SUBAPPLICATION Uebung_142_AX (* Übung zu NMEA 2000 Fast Packet senden (PGN 0x1FF00, 32 Byte) *)
  (* Standard: 61499-2; Description: Copyright (c) 2026 Meisterschulen am Ostbahnhof This program and the accompanying materials are made available under the terms of the Eclipse Public License 2.0 which is available at https://www.eclipse.org/legal/epl-2.0/ SPDX-License-Identifier: EPL-2.0 *)
  (* Version 1.0, 2026-11-17, Franz Höpfinger, Meisterschulen am Ostbahnhof, initial API and implementation and/or initial documentation *)
  PACKAGE Uebungen;
  IMPORT Uebungen::const::Uebung_120_129::Filter::ADD_ALL_PASS;
  IMPORT Uebungen::const::Uebung_120_129::Filter::FLT_ALL_PASS;
  IMPORT isobus::pgn::ADDRESS::GLOBAL_A;
  IMPORT isobus::pgn::ISOUSERHOME_e::thisMember;
  IMPORT isobus::pgn::ISO_CAN_NODE::NODE1;
  IMPORT Uebungen::const::Uebung_140_149::FastPacket::PGN_FPT_PROP_00;
  IMPORT logiBUS::io::DI::logiBUS_DI::Input_I1;
  IMPORT logiBUS::io::DI::logiBUS_DI_Events::BUTTON_SINGLE_CLICK;
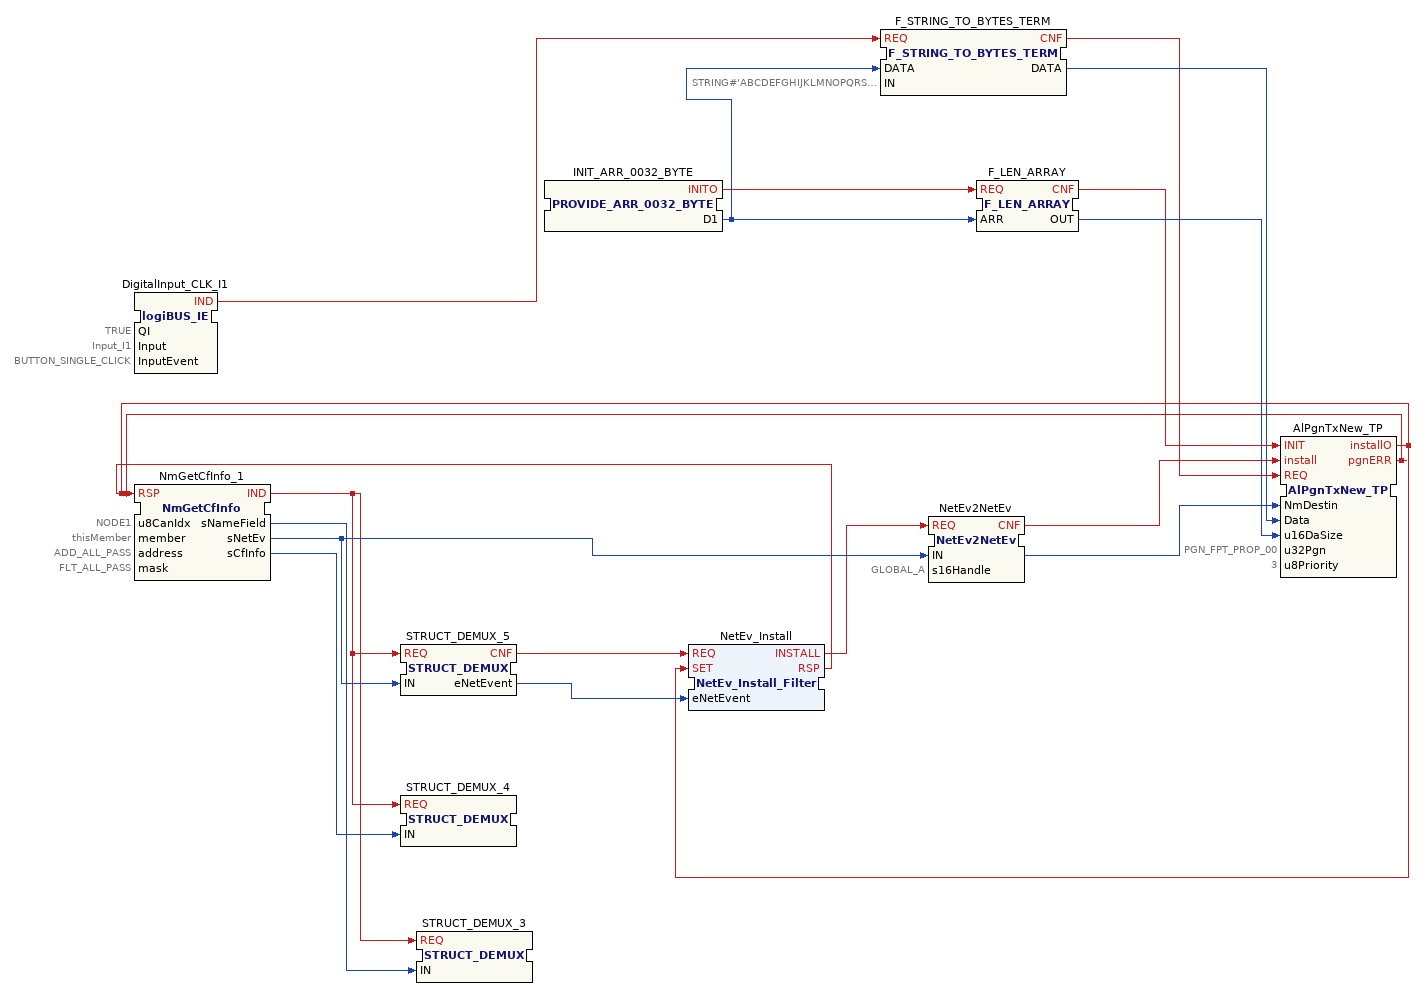
  (* NMEA 2000 Fast Packet senden: PGN 0x1FF00 (proprietär, PDU2), 32 Byte, global I1 Klick: Text A-Z 0-4 + 16#00 geht per Fast Packet (nicht ISO-TP), kein RTS/CTS. Auf dem Bus (alle mit ID 0x1FF00): Rahmen 0 = Byte0 Sequenz/Rahmenzähler, Byte1 Länge 32 (0x20), dann ABCDEF. Rahmen 1-4 = Byte0 Zähler + je 7 Daten: GHIJKLM, NOPQRST, UVWXYZ0, 1234 00 FF FF. Gegenstück: Übung 143. Firmware ab LOGIBUS 6dd74ef4 auf BEIDEN Geräten (ISO_NMEA_FPT). *)
  FBS
    STRUCT_DEMUX_3 : eclipse4diac::convert::STRUCT_DEMUX; {SET_ATTRIBUTE(StructuredType, isobus::pgn::NAMEFIELD_T)}
    NmGetCfInfo_1 : isobus::pgn::NmGetCfInfo(u8CanIdx := NODE1, member := thisMember, address := ADD_ALL_PASS, mask := FLT_ALL_PASS);
    STRUCT_DEMUX_4 : eclipse4diac::convert::STRUCT_DEMUX; {SET_ATTRIBUTE(StructuredType, isobus::pgn::CF_INFO_T)}
    STRUCT_DEMUX_5 : eclipse4diac::convert::STRUCT_DEMUX; {SET_ATTRIBUTE(StructuredType, isobus::pgn::ISONETEVENT_T)}
    NetEv2NetEv : isobus::pgn::NetEv2NetEv(s16Handle := GLOBAL_A);
    INIT_ARR_0032_BYTE : eclipse4diac::convert::providers::PROVIDE_ARR_0032_BYTE;
    F_LEN_ARRAY : eclipse4diac::utils::arrays::F_LEN_ARRAY;
    F_STRING_TO_BYTES_TERM : logiBUS::utils::dyn_arr::F_STRING_TO_BYTES_TERM(IN := STRING#'ABCDEFGHIJKLMNOPQRSTUVWXYZ01234');
    AlPgnTxNew_TP : isobus::pgn::tx::AlPgnTxNew_TP(u32Pgn := PGN_FPT_PROP_00, u8Priority := 3);
    DigitalInput_CLK_I1 : logiBUS::io::DI::logiBUS_IE(QI := TRUE, Input := Input_I1, InputEvent := BUTTON_SINGLE_CLICK);
  END_FBS
  SUBAPPS
    NetEv_Install : MyLib::sys::NetEv_Install_Filter;
  END_SUBAPPS
  EVENT_CONNECTIONS
    NmGetCfInfo_1.IND TO STRUCT_DEMUX_3.REQ;
    NmGetCfInfo_1.IND TO STRUCT_DEMUX_4.REQ;
    NmGetCfInfo_1.IND TO STRUCT_DEMUX_5.REQ;
    DigitalInput_CLK_I1.IND TO F_STRING_TO_BYTES_TERM.REQ;
    INIT_ARR_0032_BYTE.INITO TO F_LEN_ARRAY.REQ;
    F_LEN_ARRAY.CNF TO AlPgnTxNew_TP.INIT;
    NetEv2NetEv.CNF TO AlPgnTxNew_TP.install;
    F_STRING_TO_BYTES_TERM.CNF TO AlPgnTxNew_TP.REQ;
    AlPgnTxNew_TP.installO TO NmGetCfInfo_1.RSP;
    AlPgnTxNew_TP.pgnERR TO NmGetCfInfo_1.RSP;
    STRUCT_DEMUX_5.CNF TO NetEv_Install.REQ;
    NetEv_Install.INSTALL TO NetEv2NetEv.REQ;
    NetEv_Install.RSP TO NmGetCfInfo_1.RSP;
    AlPgnTxNew_TP.installO TO NetEv_Install.SET;
  END_CONNECTIONS
  DATA_CONNECTIONS
    NmGetCfInfo_1.sNameField TO STRUCT_DEMUX_3.IN;
    NmGetCfInfo_1.sNetEv TO STRUCT_DEMUX_5.IN;
    NmGetCfInfo_1.sCfInfo TO STRUCT_DEMUX_4.IN;
    NmGetCfInfo_1.sNetEv TO NetEv2NetEv.IN;
    NetEv2NetEv. TO AlPgnTxNew_TP.NmDestin;
    INIT_ARR_0032_BYTE.D1 TO F_LEN_ARRAY.ARR;
    INIT_ARR_0032_BYTE.D1 TO F_STRING_TO_BYTES_TERM.DATA;
    F_STRING_TO_BYTES_TERM.DATA TO AlPgnTxNew_TP.Data;
    F_LEN_ARRAY.OUT TO AlPgnTxNew_TP.u16DaSize;
    STRUCT_DEMUX_5.eNetEvent TO NetEv_Install.eNetEvent;
  END_CONNECTIONS
END_SUBAPPLICATION
